FUNCTION_BLOCK FB_LintTest EXTENDS FB_LintBase IMPLEMENTS I_LintItf
VAR_INPUT
END_VAR
VAR_OUTPUT
END_VAR
VAR
	nVal : INT;
	sTxt : STRING(40);
END_VAR

nVal := nVal + 1;
A_Act();

ACTION A_Act:
sTxt := 'a]]>b'; // CDATA end marker inside code
END_ACTION

METHOD PUBLIC M_Do : BOOL
M_Do := TRUE;
END_METHOD

PROPERTY PUBLIC P_Ro : INT
GET // PUBLIC
P_Ro := 1;
END_GET
END_PROPERTY

PROPERTY PUBLIC P_Val : INT
GET // PUBLIC
P_Val := nVal;
END_GET
SET // PUBLIC
nVal := P_Val;
END_SET
END_PROPERTY

END_FUNCTION_BLOCK

(* stored: Version 1.1.0.1, ProductVersion 3.1.4024.16
   POU FB_LintTest: Id {640154ed-84e6-465c-81ba-fb60f6af63e4}, SpecialFunc None
   Action A_Act: Id {7d43ebdd-86bb-4740-94ae-1ddbe750970f}
   Method M_Do: Id {f5ac9f57-167c-457b-a9c5-522abe0a7fee}
   Property P_Ro: Id {2efcd368-e92e-4201-9c00-77d6aa7999fd}
   Get Get: Id {2853db67-3245-4e9b-9cbe-74851b52738c}
   Property P_Val: Id {1da0ba76-ff51-4711-8b40-f592430ffbe3}
   Get Get: Id {25fdaa24-aa48-46a7-b470-ff71db2e5304}
   Set Set: Id {b4773b41-ea67-4819-b3a3-f76bfd5b47d9} *)
